// TIA Portal V21 export
VAR_GLOBAL   // PLC tag table "Tags_IO"
   StartButton AT %I0.0 : Bool;   // Starttaster / Start push button
   StopButton AT %I0.1 : Bool;   // Stopptaster, Öffner / Stop push button, normally closed
   LevelHigh AT %I0.2 : Bool;   // Behälterstand hoch / Tank level high
   SelectorInputs AT %IB1 : Byte;   // Eingänge Betriebsartenwahlschalter / Mode selector inputs
   FlowRaw AT %IW2 : Word;   // Rohwert Durchfluss / Raw flow value
   ConveyorRun AT %Q0.0 : Bool;   // Fördermotor ein / Conveyor motor on
   ValveOpen AT %Q0.1 : Bool;   // Füllventil auf / Filling valve open
   LampOutputs AT %QB1 : Byte;   // Signalleuchten / Signal lamps
   SpeedOutput AT %QW2 : Word;   // Drehzahlsollwert an den Antrieb / Speed setpoint to the drive
END_VAR
